Universal Robots URScript: program3.script

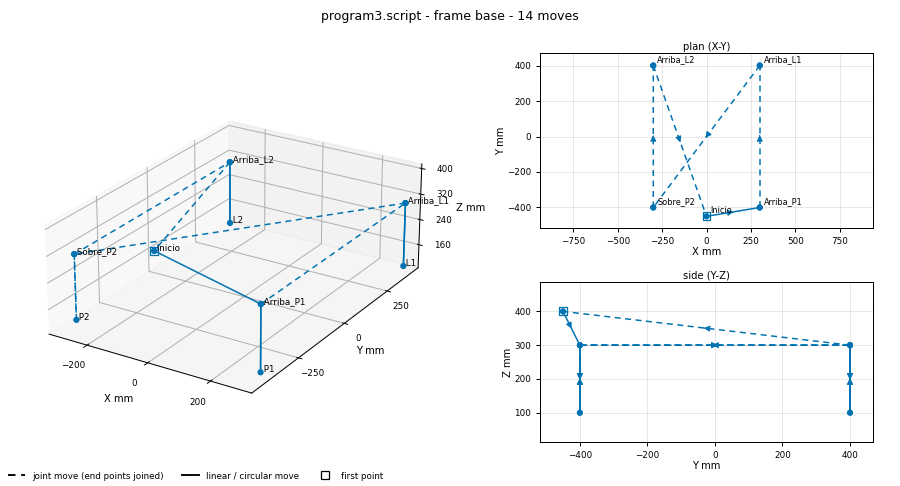
[picture p0: tool path of program3.script in frame base, 14 of 14 moves have a stored position in this frame; points joined in program order, loops and branches not executed]
def program3():
  set_safety_mode_transition_hardness(1)
  set_tcp(p[0.0,0.0,0.0,0.0,0.0,0.0])
  set_payload(0.0)
  set_gravity([0.0, 0.0, 9.82])
  set_standard_analog_input_domain(0, 1)
  set_standard_analog_input_domain(1, 1)
  set_tool_analog_input_domain(0, 1)
  set_tool_analog_input_domain(1, 1)
  set_analog_outputdomain(0, 0)
  set_analog_outputdomain(1, 0)
  set_input_actions_to_default()
  step_count_32e24061_6999_48a6_b80b_3f88d94f556b = 0.0
  thread Step_Counter_Thread_853c1897_7aa5_40e5_bd8d_e01aeb857cb3():
    while (True):
      step_count_32e24061_6999_48a6_b80b_3f88d94f556b = step_count_32e24061_6999_48a6_b80b_3f88d94f556b + 1.0
      sync()
    end
  end
  run Step_Counter_Thread_853c1897_7aa5_40e5_bd8d_e01aeb857cb3()
  set_tool_voltage(0)
  # begin: URCap Installation Node
  #   Source: External Control, 1.0.5, FZI Research Center for Information Technology
  #   Type: External Control
  # end: URCap Installation Node
  while (True):
    $ 1 "Robot Program"
    $ 2 "MoveJ"
    $ 3 "Inicio" "breakAfter"
    movej(get_inverse_kin(p[.000000003418, -.449999953698, .400000040186, -3.141185387045, .000000412671, .000000636370], qnear=[1.3258157968521118, -1.686899487172262, 1.7607979774475098, -1.6442998091327112, -1.5708954969989222, 2.8966124057769775]), a=1.3962634015954636, v=1.0471975511965976)
    $ 4 "MoveL"
    $ 5 "Arriba_P1" "breakAfter"
    movel(p[.300000000000, -.400000000000, .300000000000, -3.141185387046, .000000412671, .000000636369], a=1.2, v=0.25)
    $ 6 "P1" "breakAfter"
    movel(p[.300000000000, -.400000000000, .100000000000, -3.141185387046, .000000000000, .000000000000], a=1.2, v=0.25)
    $ 7 "Set DO[1]=On"
    set_standard_digital_out(1, True)
    set_payload(1.0)
    $ 8 "Wait: 0.5"
    sleep(0.5)
    $ 9 "MoveL"
    $ 10 "Subir_P1" "breakAfter"
    movel(p[.300000000000, -.400000000000, .300000000000, -3.141185387046, .000000000000, .000000000000], a=1.2, v=0.25)
    $ 11 "Wait: 1.0"
    sleep(1.0)
    $ 12 "MoveJ"
    $ 13 "Arriba_L1" "breakAfter"
    movej(get_inverse_kin(p[.300000000000, .400000000000, .300000000000, -3.141185387046, .000000000000, .000000000000], qnear=[3.8487635350581386, -1.5152013940703055, 1.8563295772739679, -1.9121891054490625, -1.570486721364162, 5.419559902608085]), a=1.3962634015954636, v=1.0471975511965976)
    $ 14 "MoveL"
    $ 15 "L1" "breakAfter"
    movel(p[.300000000000, .400000000000, .100000000000, -3.141185387046, .000000000000, .000000000000], a=1.2, v=0.25)
    $ 16 "Set DO[1]=Off"
    set_standard_digital_out(1, False)
    set_payload(0.0)
    $ 17 "Wait: 0.5"
    sleep(0.5)
    $ 18 "MoveL"
    $ 19 "Subir_L1" "breakAfter"
    movel(p[.300000000000, .400000000000, .300000000000, -3.141185387046, .000000000000, .000000000000], a=1.2, v=0.25)
    $ 20 "MoveJ"
    $ 21 "Sobre_P2" "breakAfter"
    movej(get_inverse_kin(p[-.300017425944, -.399967031817, .299973586294, -3.141100507342, -.000000095361, -.000060560188], qnear=[0.7072074129081024, -1.5151203236562776, 1.8561576594959694, -1.9114845967841896, -1.5711453926452954, 2.2780037397029993]), a=1.3962634015954636, v=1.0471975511965976)
    $ 22 "MoveJ"
    $ 23 "P2" "breakAfter"
    movej(get_inverse_kin(p[-.300015527182, -.399965408919, .099956561067, -3.141100507342, -.000000095361, -.000060560189], qnear=[0.7072074129081024, -1.2168435544904466, 2.1097539998107453, -2.4633577062647967, -1.5711453926452954, 2.2780037397029993]), a=1.3962634015954636, v=1.0471975511965976)
    $ 24 "Set DO[1]=On"
    set_standard_digital_out(1, True)
    set_payload(1.0)
    $ 25 "Wait: 0.5"
    sleep(0.5)
    $ 26 "MoveJ"
    $ 27 "Subir_P2" "breakAfter"
    movej(get_inverse_kin(p[-.300017425944, -.399967031817, .299973586294, -3.141100507341, -.000000095361, -.000060560188], qnear=[0.7072074129081024, -1.5151203236562776, 1.8561576594959694, -1.9114845967841896, -1.5711453926452954, 2.2780037397029993]), a=1.3962634015954636, v=1.0471975511965976)
    $ 28 "Wait: 1.0"
    sleep(1.0)
    $ 29 "MoveJ"
    $ 30 "Arriba_L2" "breakAfter"
    movej(get_inverse_kin(p[-.299958791196, .399992870398, .300007996726, 3.141482059736, .000000076039, .000679639003], qnear=[-1.1473794502610721, -1.5151908478860783, 1.8561576594959694, -1.9114845967841896, -1.5711453926452954, 0.42341687653382437]), a=1.3962634015954636, v=1.0471975511965976)
    $ 31 "MoveL"
    $ 32 "L2" "breakAfter"
    movel(p[-.299963931488, .400004276205, .099950247894, 3.141405955254, .000000098917, .000733486799], a=1.2, v=0.25)
    $ 33 "Set DO[1]=Off"
    set_standard_digital_out(1, False)
    set_payload(0.0)
    $ 34 "Wait: 0.5"
    sleep(0.5)
    $ 35 "MoveL"
    $ 36 "Subir_L2" "breakAfter"
    movel(p[-.299958791196, .399992870398, .300007996726, 3.141482059736, .000000076039, .000679639003], a=1.2, v=0.25)
    $ 37 "MoveJ"
    $ 38 "Fin" "breakAfter"
    movej(get_inverse_kin(p[.000000000000, -.450000000000, .400000000000, -3.141185307180, .000000000000, .000000000000], qnear=[1.3258157445438208, -1.686899352753934, 1.7607979201646433, -1.6442997105343231, -1.5708951233618098, 2.89661209065496]), a=1.3962634015954636, v=1.0471975511965976)
    $ 39 "Wait DI[0]=HI"
    while (get_standard_digital_in(0) == False):
      sync()
    end
  end
end
